FUNCTION_BLOCK PhasesOff (* Emergencia: indica, para ate 7 fases, se a fase esta parada (equipamentos desligados) *)
  (* Standard: 61499-2 *)
  (* Version 1.0, 30/10/2026, Hidryco, Hidryco, 1.0: Off = estado fora de Starting/Running/Stopping/Aborting (Ready, Aborted, Interlocked ou vazio). Usado para o passo da emergencia so terminar com a fase parada. *)
  PACKAGE SE.Nereda;
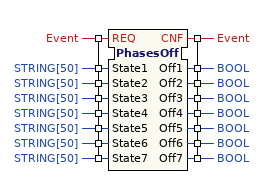
  EVENT_INPUT
    REQ WITH State1, State2, State3, State4, State5, State6, State7; (* Mudanca de estado de alguma fase *)
  END_EVENT
  EVENT_OUTPUT
    CNF WITH Off1, Off2, Off3, Off4, Off5, Off6, Off7;
  END_EVENT
  VAR_INPUT
    State1 : STRING[50]; (* Estado da fase 1 (Phase.State); vazio = sem fase *)
    State2 : STRING[50]; (* Estado da fase 2 (Phase.State); vazio = sem fase *)
    State3 : STRING[50]; (* Estado da fase 3 (Phase.State); vazio = sem fase *)
    State4 : STRING[50]; (* Estado da fase 4 (Phase.State); vazio = sem fase *)
    State5 : STRING[50]; (* Estado da fase 5 (Phase.State); vazio = sem fase *)
    State6 : STRING[50]; (* Estado da fase 6 (Phase.State); vazio = sem fase *)
    State7 : STRING[50]; (* Estado da fase 7 (Phase.State); vazio = sem fase *)
  END_VAR
  VAR_OUTPUT
    Off1 : BOOL := TRUE; (* Fase 1 parada (nao esta em Starting/Running/Stopping/Aborting) *)
    Off2 : BOOL := TRUE; (* Fase 2 parada (nao esta em Starting/Running/Stopping/Aborting) *)
    Off3 : BOOL := TRUE; (* Fase 3 parada (nao esta em Starting/Running/Stopping/Aborting) *)
    Off4 : BOOL := TRUE; (* Fase 4 parada (nao esta em Starting/Running/Stopping/Aborting) *)
    Off5 : BOOL := TRUE; (* Fase 5 parada (nao esta em Starting/Running/Stopping/Aborting) *)
    Off6 : BOOL := TRUE; (* Fase 6 parada (nao esta em Starting/Running/Stopping/Aborting) *)
    Off7 : BOOL := TRUE; (* Fase 7 parada (nao esta em Starting/Running/Stopping/Aborting) *)
  END_VAR
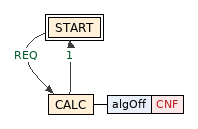
  EC_STATES
    START; (* Initial State *)
    CALC : algOff -> CNF;
  END_STATES
  EC_TRANSITIONS
    START TO CALC := REQ;
    CALC TO START := 1;
  END_TRANSITIONS
  ALGORITHM algOff IN ST:
Off1 := NOT (State1 = 'Starting' OR State1 = 'Running' OR State1 = 'Stopping' OR State1 = 'Aborting');
Off2 := NOT (State2 = 'Starting' OR State2 = 'Running' OR State2 = 'Stopping' OR State2 = 'Aborting');
Off3 := NOT (State3 = 'Starting' OR State3 = 'Running' OR State3 = 'Stopping' OR State3 = 'Aborting');
Off4 := NOT (State4 = 'Starting' OR State4 = 'Running' OR State4 = 'Stopping' OR State4 = 'Aborting');
Off5 := NOT (State5 = 'Starting' OR State5 = 'Running' OR State5 = 'Stopping' OR State5 = 'Aborting');
Off6 := NOT (State6 = 'Starting' OR State6 = 'Running' OR State6 = 'Stopping' OR State6 = 'Aborting');
Off7 := NOT (State7 = 'Starting' OR State7 = 'Running' OR State7 = 'Stopping' OR State7 = 'Aborting');
  END_ALGORITHM
END_FUNCTION_BLOCK
